RESOURCE RES0 : EMB_RES_ECO
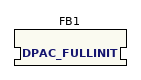
  FBS
    FB1 : DPAC_FULLINIT;
  END_FBS
END_RESOURCE
